Fanuc KAREL source: KO00010.KL

PROGRAM KO00010
%NOLOCKGROUP
VAR
  P1: XYZWPR
  P2: XYZWPR
  P3: XYZWPR
  OUT: XYZWPR
BEGIN
  OUT = FRAME(P1, P2, P3)
END KO00010
